(* Logix 5000 project; controller ViciOne vendor 1 type 14 code 196 rev 36.11; software revision 36.00 *)

TASK MainTask (continuous, watchdog 500 ms) : MainProgram

MODULES
   Local : vendor 1 type 14 code 196 (5069 0, rev 36.11)
      INPUT : 5069-IB16 (5069 1, rev 2.16, StandardDataDriven RPI 5 ms)
      OUTPUT : 5069-OB16 (5069 2, rev 3.13, StandardDataDriven RPI 5 ms)
END_MODULES

TYPE STRING_20 :
STRUCT
   LEN : DINT;
   DATA : SINT[20];
END_STRUCT
END_TYPE

TYPE UDT_Inner :
STRUCT
   BoolTag : BOOL;
   RealTag : REAL;
   IntArray : INT[10];
   StringTag : STRING;
END_STRUCT
END_TYPE

TYPE UDT_Outer :
STRUCT
   BoolTag : BOOL;
   BoolNeighbour : BOOL;
   DIntTag : DINT;
   StringTag : STRING;
   String20 : STRING_20;
   DIntArray : DINT[10];
   BoolArray : BOOL[32];
   TimerTag : TIMER;
   TimerArray : TIMER[10];
   CounterTag : COUNTER;
   InnerUdt : UDT_Inner;
END_STRUCT
END_TYPE

VAR_GLOBAL   (* controller tags *)
   BoolArrayControllerTag : BOOL[32] := ([0] := 1, [1] := 1, [7] := 1, [8] := 1, [15] := 1, [16] := 1, [30] := 1, [31] := 1);
   BoolControllerTag : BOOL;
   CounterControllerTag : COUNTER := (PRE := 500);
   DIntArrayControllerTag : DINT[10] := ([1] := 1, [2] := -1, [3] := 123456, [4] := -2147483648, [5] := 2147483647, [6] := 10, [7] := 20, [8] := 30, [9] := 40);
   DIntControllerTag : DINT := 123456;
   DIntTag : DINT := 1111;   // Provisioned under this name in both scopes, so the program tag shadows the controller tag.
   IntArrayControllerTag : INT[10] := ([1] := 1, [2] := -1, [3] := 4711, [4] := -32768, [5] := 32767, [6] := 10, [7] := 20, [8] := 30, [9] := 40);
   IntControllerTag : INT := -1;
   LIntArrayControllerTag : LINT[10] := ([1] := 1, [2] := -1, [3] := 1234567890123, [4] := -9223372036854775808, [5] := 9223372036854775807, [6] := 10, [7] := 20, [8] := 30, [9] := 40);
   LIntControllerTag : LINT := 9223372036854775807;
   LRealArrayControllerTag : LREAL[10] := ([1] := 1.0, [2] := -1.0, [3] := 3.141592653589793, [4] := -1.7976931348623157e+308, [5] := 1.7976931348623157e+308, [6] := 10.5, [7] := -20.25, [8] := 30.75, [9] := 40.0);
   LRealControllerTag : LREAL := -1.7976931348623157e+308;
   RealArrayControllerTag : REAL[10] := ([1] := 1.0, [2] := -1.0, [3] := 3.14159, [6] := 10.5, [7] := -20.25, [8] := 30.75, [9] := 40.0);
   RealControllerTag : REAL;
   SIntArrayControllerTag : SINT[10] := ([1] := 1, [2] := -1, [3] := 42, [4] := -128, [5] := 127, [6] := 10, [7] := 20, [8] := 30, [9] := 40);
   SIntControllerTag : SINT := 42;
   String20ControllerTag : STRING_20 := 'XXXXXXXXXXXXXXXXXXXX';
   StringControllerTag : STRING := 'XXXXXXXXXXXXXXXXXXXXXXXXXXXXXXXXXXXXXXXXXXXXXXXXXXXXXXXXXXXXXXXXXXXXXXXXXXXXXXXXXX';
   TimerArrayControllerTag : TIMER[10] := ([3].ACC := 1234);
   TimerControllerTag : TIMER := (PRE := 5000, ACC := 1234);
   UDIntArrayControllerTag : UDINT[10] := ([3] := 4000000000);
   UDIntControllerTag : UDINT := 2147483648;
   UdtControllerTag : UDT_Outer := (BoolNeighbour := 1, DIntTag := 123456, StringTag := 'Hello World', String20 := 'XXXXXXXXXXXXXXXXXXXX', DIntArray[0] := -2147483648, DIntArray[1] := -1, DIntArray[3] := 1, DIntArray[4] := 123456, DIntArray[5] := 5, DIntArray[6] := 6, DIntArray[7] := 7, DIntArray[8] := 8, DIntArray[9] := 2147483647, BoolArray[0] := 1, BoolArray[1] := 1, BoolArray[7] := 1, BoolArray[8] := 1, BoolArray[15] := 1, BoolArray[16] := 1, BoolArray[30] := 1, BoolArray[31] := 1, TimerTag.PRE := 5000, TimerTag.ACC := 1234, TimerArray[3].ACC := 1234, CounterTag.ACC := -1234, InnerUdt.BoolTag := 1, InnerUdt.RealTag := 123.456, InnerUdt.IntArray[3] := 4711, InnerUdt.StringTag := 'Nested');
   UIntArrayControllerTag : UINT[10] := ([3] := 50000);
   UIntControllerTag : UINT := 65535;
   ULIntArrayControllerTag : ULINT[10] := ([3] := 18446744073709551614);
   ULIntControllerTag : ULINT;
   USIntArrayControllerTag : USINT[10] := ([3] := 200);
   USIntControllerTag : USINT := 255;
END_VAR

PROGRAM MainProgram   (* main routine MainRoutine *)
// Integration-suite tags. Every tag here, and every controller tag, is written by the test suites; no instruction may use one.
VAR
   BoolArrayProgramTag : BOOL[32] := ([0] := 1, [1] := 1, [7] := 1, [8] := 1, [15] := 1, [16] := 1, [30] := 1, [31] := 1);
   BoolProgramTag : BOOL;
   Counter : COUNTER;   // Mirrors the L32E, for the CompactLogix5X70 suite. The suite reads Counter.PRE.
   CounterProgramTag : COUNTER := (PRE := 500, ACC := 1234);
   DIntArrayProgramTag : DINT[10] := ([1] := 1, [2] := -1, [3] := 123456, [4] := -2147483648, [5] := 2147483647, [6] := 10, [7] := 20, [8] := 30, [9] := 40);
   DIntProgramTag : DINT := 123456;
   DIntTag : DINT := 2222;   // Provisioned under this name in both scopes, so the program tag shadows the controller tag.
   IntArrayProgramTag : INT[10] := ([1] := 1, [2] := -1, [3] := 4711, [4] := -32768, [5] := 32767, [6] := 10, [7] := 20, [8] := 30, [9] := 40);
   IntProgramTag : INT := -1;
   LIntArrayProgramTag : LINT[10] := ([1] := 1, [2] := -1, [3] := 1234567890123, [4] := -9223372036854775808, [5] := 9223372036854775807, [6] := 10, [7] := 20, [8] := 30, [9] := 40);
   LIntProgramTag : LINT := -9223372036854775808;
   LRealArrayProgramTag : LREAL[10] := ([3] := 3.141592653589793);
   LRealProgramTag : LREAL;
   RealArrayProgramTag : REAL[10] := ([3] := 3.14159);
   RealProgramTag : REAL;
   SIntArrayProgramTag : SINT[10] := ([1] := 1, [2] := -1, [3] := 42, [4] := -128, [5] := 127, [6] := 10, [7] := 20, [8] := 30, [9] := 40);
   SIntProgramTag : SINT := 127;
   String20ProgramTag : STRING_20 := 'XXXXXXXXXXXXXXXXXXXX';
   StringProgramTag : STRING := 'Hello World';
   strValue1 : STRING;   // Mirrors the L32E, for the CompactLogix5X70 suite.
   TimerArrayProgramTag : TIMER[10] := ([3].ACC := 1234);
   TimerProgramTag : TIMER := (PRE := 5000, ACC := 55);
   UDIntArrayProgramTag : UDINT[10] := ([1] := 1, [2] := 123456, [3] := 2147483648, [4] := 4000000000, [5] := 4294967295, [6] := 10, [7] := 20, [8] := 30, [9] := 40);
   UDIntProgramTag : UDINT := 2147483648;
   UdtProgramTag : UDT_Outer := (BoolTag := 1, DIntTag := 33, StringTag := 'Hello World', String20 := 'XXXXXXXXXXXXXXXXXXXX', DIntArray[3] := 123456, BoolArray[0] := 1, BoolArray[1] := 1, BoolArray[7] := 1, BoolArray[8] := 1, BoolArray[15] := 1, BoolArray[16] := 1, BoolArray[30] := 1, BoolArray[31] := 1, TimerTag.PRE := 5000, TimerTag.ACC := 1234, TimerArray[3].ACC := 1234, CounterTag.ACC := -1234, InnerUdt.RealTag := 44.5, InnerUdt.IntArray[3] := 4711, InnerUdt.StringTag := 'Nested');
   UIntArrayProgramTag : UINT[10] := ([1] := 1, [2] := 4242, [3] := 32768, [4] := 50000, [5] := 65535, [6] := 10, [7] := 20, [8] := 30, [9] := 40);
   UIntProgramTag : UINT := 65535;
   ULIntArrayProgramTag : ULINT[10] := ([1] := 1, [2] := 1234567890123, [3] := 9223372036854775808, [4] := 18446744073709551614, [5] := 18446744073709551615, [6] := 10, [7] := 20, [8] := 30, [9] := 40);
   ULIntProgramTag : ULINT := 1234567890123;
   USIntArrayProgramTag : USINT[10] := ([1] := 1, [2] := 42, [3] := 128, [4] := 200, [5] := 255, [6] := 10, [7] := 20, [8] := 30, [9] := 40);
   USIntProgramTag : USINT := 42;
END_VAR

ROUTINE MainRoutine   (* ladder *)
   0: NOP();
END_ROUTINE
END_PROGRAM
